FUNCTION_BLOCK SimulatedValve IMPLEMENTS I_FillValve, I_Cyclic
VAR
    _Name         : STRING(32);
    _Clock        : I_Clock;
    _TravelTime   : LTIME;
    _IsCommanded  : BOOL;              // TRUE: open requested
    _IsStuck      : BOOL;
    _IsAtOpen     : BOOL;
    _IsAtClosed   : BOOL := TRUE;
    _MoveStart    : LTIME;
    _IsMoving     : BOOL;
    _IsConfigured : BOOL;
END_VAR
(*
    SimulatedValve

    Stands in for a valve with position feedback. Reaches the commanded
    position after TravelTime, with neither end reported while it moves.
    SetStuck() makes it stop answering commands, as a sticking valve does.
    Has no I/O.
*)

METHOD FB_init : BOOL
VAR_INPUT
    bInitRetains : BOOL;
    bInCopyCode  : BOOL;
    Name         : STRING(32);
    Clock        : I_Clock;
    TravelTime   : LTIME;
END_VAR
_Name := Name;
_Clock := Clock;
_TravelTime := TravelTime;
_IsConfigured := Clock <> 0;
END_METHOD

METHOD PUBLIC Open
_IsCommanded := TRUE;
END_METHOD

METHOD PUBLIC Close
_IsCommanded := FALSE;
END_METHOD

METHOD PUBLIC SetStuck
VAR_INPUT
    IsStuck : BOOL;
END_VAR
_IsStuck := IsStuck;
END_METHOD

METHOD PUBLIC CyclicLogic
IF NOT _IsConfigured OR _IsStuck THEN
    RETURN;
END_IF
IF _IsCommanded <> _IsAtOpen AND NOT _IsMoving THEN
    _IsMoving := TRUE;                 // a new command: leave the end position
    _MoveStart := _Clock.Now;
    _IsAtOpen := FALSE;
    _IsAtClosed := FALSE;
END_IF
IF _IsMoving AND_THEN _Clock.Now - _MoveStart >= _TravelTime THEN
    _IsMoving := FALSE;
    _IsAtOpen := _IsCommanded;
    _IsAtClosed := NOT _IsCommanded;
END_IF
END_METHOD

PROPERTY PUBLIC IsOpen : BOOL
GET
IsOpen := _IsAtOpen;
END_GET
END_PROPERTY

PROPERTY PUBLIC IsClosed : BOOL
GET
IsClosed := _IsAtClosed;
END_GET
END_PROPERTY

PROPERTY PUBLIC Name : STRING
GET
Name := _Name;
END_GET
END_PROPERTY

PROPERTY PUBLIC HasFault : BOOL
GET
HasFault := NOT _IsConfigured;
END_GET
END_PROPERTY

PROPERTY PUBLIC FaultText : STRING
GET
FaultText := SEL(_IsConfigured, 'Simulated valve has no clock', '');
END_GET
END_PROPERTY

END_FUNCTION_BLOCK

(* stored: Version 1.1.0.1, ProductVersion 3.1.4026.0
   POU SimulatedValve: Id {50001f74-fdd6-4023-9443-28f93956bd61}, SpecialFunc None
   Folder I_FillValve: Id {39ace360-a19f-444c-8b46-74e312015064}
   Folder I_Diagnosable: Id {6bdeec5e-a873-4a84-8a60-1505c70f6ac2}
   Folder I_Cyclic: Id {1adbcab9-caf9-4d33-a28a-fb94d523ff33}
   Method FB_init: Id {573dd73e-ff25-408d-830d-627946ceb760}
   Method Open: Id {be3bd5c9-a304-4e1d-b694-5ba0ebb77cc5}
   Method Close: Id {8ef05bd0-9ef9-495b-91aa-6b4d2cb1211c}
   Method SetStuck: Id {9780cfa5-ae8d-4c18-bc8a-734a5e7d0b85}
   Method CyclicLogic: Id {d169821f-5edd-4d6b-b58a-f54406e4d385}
   Property IsOpen: Id {401f1036-a01d-4bbc-a6f2-b8c9aae2efab}
   Get Get: Id {20edcc6d-c550-4669-aea1-784ba0aad3ab}
   Property IsClosed: Id {82ebd267-6267-4dcd-b2b9-b2714623ed67}
   Get Get: Id {6e603605-20f8-4a79-a181-526ba2782219}
   Property Name: Id {47186d54-ed5b-4137-ab87-0163d556528c}
   Get Get: Id {077bf48f-4d56-42cc-a599-a68436ebbd4a}
   Property HasFault: Id {53cdd4eb-11e2-4542-9190-0a61c515d2fc}
   Get Get: Id {3b6a8322-167e-4cc7-9394-9ca87ee0520d}
   Property FaultText: Id {de07335c-7968-4fa5-a76f-1c5b7c1a3943}
   Get Get: Id {765de1ea-0d49-4ee8-be7f-19ac3c5e2ef9} *)
